(* IEC 61131-3 sources: PLCHaT-dataset/benchmark_mutated/222_MaterialMixing/mutation_3/plc_st_files, 1 file *)

(* ---- 222_MaterialMixing.st ---- *)
FUNCTION_BLOCK MaterialMixing
VAR_INPUT
estop : BOOL; (* Emergency Stop Signal, FALSE: Emergency stop triggered, TRUE: No emergency stop triggered *)
opeMode : BOOL; (* Operation Mode, FALSE: Manual Operation Mode, TRUE: Automatic Operation Mode *)
valveAStart : BOOL; (* Valve A Start Button *)
valveBStart : BOOL; (* Valve B Start Button *)
valveCStart : BOOL; (* Valve C Start Button *)
valveDStart : BOOL; (* Valve D Start Button *)
mixMotorStart : BOOL; (* Mixing Motor Start Button *)
autoStart : BOOL; (* Automatic Start Button *)
processMode : BOOL; (* Process Mode *)
levelSensor : INT; (* Liquid Level Sensor, unit cm *)
END_VAR

VAR_OUTPUT
valveARun : BOOL; (* Valve A Run Command *)
valveBRun : BOOL; (* Valve B Run Command *)
valveCRun : BOOL; (* Valve C Run Command *)
valveDRun : BOOL; (* Valve D Run Command *)
mixMotorRun : BOOL; (* Mixing Motor Run Command *)
END_VAR

VAR
previousValveAStart : BOOL := FALSE;
previousValveBStart : BOOL := FALSE;
previousValveCStart : BOOL := FALSE;
previousValveDStart : BOOL := FALSE;
previousMixMotorStart : BOOL := FALSE;
previousAutoStart : BOOL := FALSE;
autoStep : INT := 0; (* Sequence step variable for automatic mode *)
mixMotorComplete : BOOL; (* Mixing Complete Signal *)

(* Temporary variables for rising edge detection - using VAR for calculation *)
valveA_RE : BOOL;
valveB_RE : BOOL;
valveC_RE : BOOL;
valveD_RE : BOOL;
mixMotor_RE : BOOL;
autoStart_RE : BOOL;
END_VAR

(* Implementation of MaterialMixing Function Block *)

(* --- 1. Emergency Stop Logic --- *)
IF NOT estop THEN
    (* Immediate stop all equipment and reset sequence *)
    valveARun := FALSE;
    valveBRun := FALSE;
    valveCRun := FALSE;
    valveDRun := FALSE;
    mixMotorRun := FALSE;
    autoStep := 0;
ELSE
    (* --- 2. Operation Mode Selection --- *)
    IF NOT opeMode THEN
        (* --- 2.1. Manual Operation Mode (opeMode = FALSE) --- *)

        autoStep := 0;

        (* Calculate Rising Edges (RE) for Manual Toggle *)
        valveA_RE := valveAStart AND NOT previousValveAStart;
        valveB_RE := valveBStart AND NOT previousValveBStart;
        valveC_RE := valveCStart AND NOT previousValveCStart;
        valveD_RE := valveDStart AND NOT previousValveDStart;
        mixMotor_RE := mixMotorStart AND NOT previousMixMotorStart;

        (* Toggle Logic on Rising Edge *)
        IF valveA_RE THEN valveARun := NOT valveARun; END_IF;
        IF valveB_RE THEN valveBRun := NOT valveBRun; END_IF;
        IF valveC_RE THEN valveCRun := NOT valveCRun; END_IF;
        IF valveD_RE THEN valveDRun := NOT valveDRun; END_IF;
        IF mixMotor_RE THEN mixMotorRun := NOT mixMotorRun; END_IF;

    ELSE
        (* --- 2.2. Automatic Operation Mode (opeMode = TRUE) --- *)

        autoStart_RE := autoStart AND NOT previousAutoStart;

        (* Reset all outputs at the beginning of the auto mode cycle *)
        valveARun := FALSE;
        valveBRun := FALSE;
        valveCRun := FALSE;
        valveDRun := FALSE;
        mixMotorRun := FALSE;

        (* --- MUTATION: Decouple level sensor from state transition logic --- *)
        (* The original logic pre-emptively adjusts autoStep based on sensor readings, *)
        (* bypassing the intended sequential state machine. This mutation removes that coupling. *)
        IF autoStep < 50 THEN (* Only applies during the filling stages *)
            (* Level sensor readings are now ignored for state advancement. *)
            (* The system must progress solely via the CASE state machine below. *)
            autoStep := autoStep;
        END_IF;

        (* --- State Machine Logic (using potentially adjusted autoStep) --- *)
        CASE autoStep OF
            0: (* Idle / Initial State *)
                IF autoStart_RE THEN
                    autoStep := 10; (* Start the process *)
                END_IF;

            10: (* Step 1: Fill A *)
                IF levelSensor >= 50 THEN
                    autoStep := 20; (* Transition: Close A, Open B *)
                    valveBRun := TRUE;  (* Immediate output change to ensure transition is complete in 1 cycle *)
                    valveARun := FALSE; (* Immediate output change *)
                ELSE
                    valveARun := TRUE;
                END_IF;

            20: (* Step 2: Fill B *)
                IF levelSensor >= 80 THEN
                    autoStep := 30; (* Transition: Close B, Check Process Mode *)
                    valveBRun := FALSE; (* Immediate output change *)
                ELSE
                    valveBRun := TRUE;
                END_IF;

            30: (* Step 3: Close Valve B, Check Process Mode *)
                IF NOT processMode THEN
                    valveCRun := FALSE;
                    autoStep := 50; (* Transition to Mixing (Mode FALSE) *)
                ELSE
                    valveCRun := TRUE;
                    autoStep := 40; (* Transition to Fill C (Mode TRUE) *)
                END_IF;

            40: (* Step 4: Process Mode TRUE: Fill C *)
                IF levelSensor >= 100 THEN
                    valveCRun := FALSE;
                    autoStep := 50; (* Transition to Mixing *)
                ELSE
                    valveCRun := TRUE;
                END_IF;

            50: (* Step 5: Start Mixing Motor *)
                IF mixMotorComplete THEN
                    mixMotorRun := FALSE; (* Stop motor *)
                    autoStep := 60; (* Transition to Delivery *)
                ELSE
                    mixMotorRun := TRUE;
                END_IF;

            60: (* Step 6: Open Valve D - Process End *)
                valveDRun := TRUE;
                IF NOT autoStart THEN
                    autoStep := 0;
                END_IF;

            ELSE
                autoStep := 0; (* Failsafe to idle state *)
        END_CASE;

    END_IF;

    (* --- 3. Update Previous Values for Next Scan Cycle --- *)
    previousValveAStart := valveAStart;
    previousValveBStart := valveBStart;
    previousValveCStart := valveCStart;
    previousValveDStart := valveDStart;
    previousMixMotorStart := mixMotorStart;
    previousAutoStart := autoStart;

END_IF;
END_FUNCTION_BLOCK
